PROGRAM main
  VAR
    S1 AT %IX0.0  : BOOL; (* abrir, NA *)
    S2 AT %IX0.1  : BOOL; (* cerrar, NA *)
    S0 AT %IX0.2  : BOOL; (* parada, NC: TRUE sin pulsar *)
    B1 AT %IX0.3  : BOOL; (* final: portón abierto *)
    B2 AT %IX0.4  : BOOL; (* final: portón cerrado *)
    B3 AT %IX0.5  : BOOL; (* barrera: obstáculo en el paso *)
    KM1 AT %QX0.0 : BOOL; (* motor: abrir *)
    KM2 AT %QX0.1 : BOOL; (* motor: cerrar *)
    H1 AT %QX0.2  : BOOL; (* baliza de movimiento *)
    ETAPA         : INT; (* 0 parado, 1 abriendo, 2 cerrando *)
    E0            : BOOL; (* ETAPA = 0 *)
    E1            : BOOL; (* ETAPA = 1 *)
    E2            : BOOL; (* ETAPA = 2 *)
  END_VAR
  VAR  (* added by the conversion: wires and edge detectors of the diagram *)
    _EQ1_OUT : BOOL;
    _EQ5_OUT : BOOL;
    _EQ9_OUT : BOOL;
    _NOT17_OUT : BOOL;
    _AND14_OUT : BOOL;
    _SEL13_OUT : INT;
    _NOT26_OUT : BOOL;
    _AND23_OUT : BOOL;
    _SEL22_OUT : INT;
    _AND32_OUT : BOOL;
    _SEL31_OUT : INT;
    _AND39_OUT : BOOL;
    _SEL38_OUT : INT;
    _AND46_OUT : BOOL;
    _SEL45_OUT : INT;
    _NOT53_OUT : BOOL;
    _SEL52_OUT : INT;
    _NOT62_OUT : BOOL;
  END_VAR

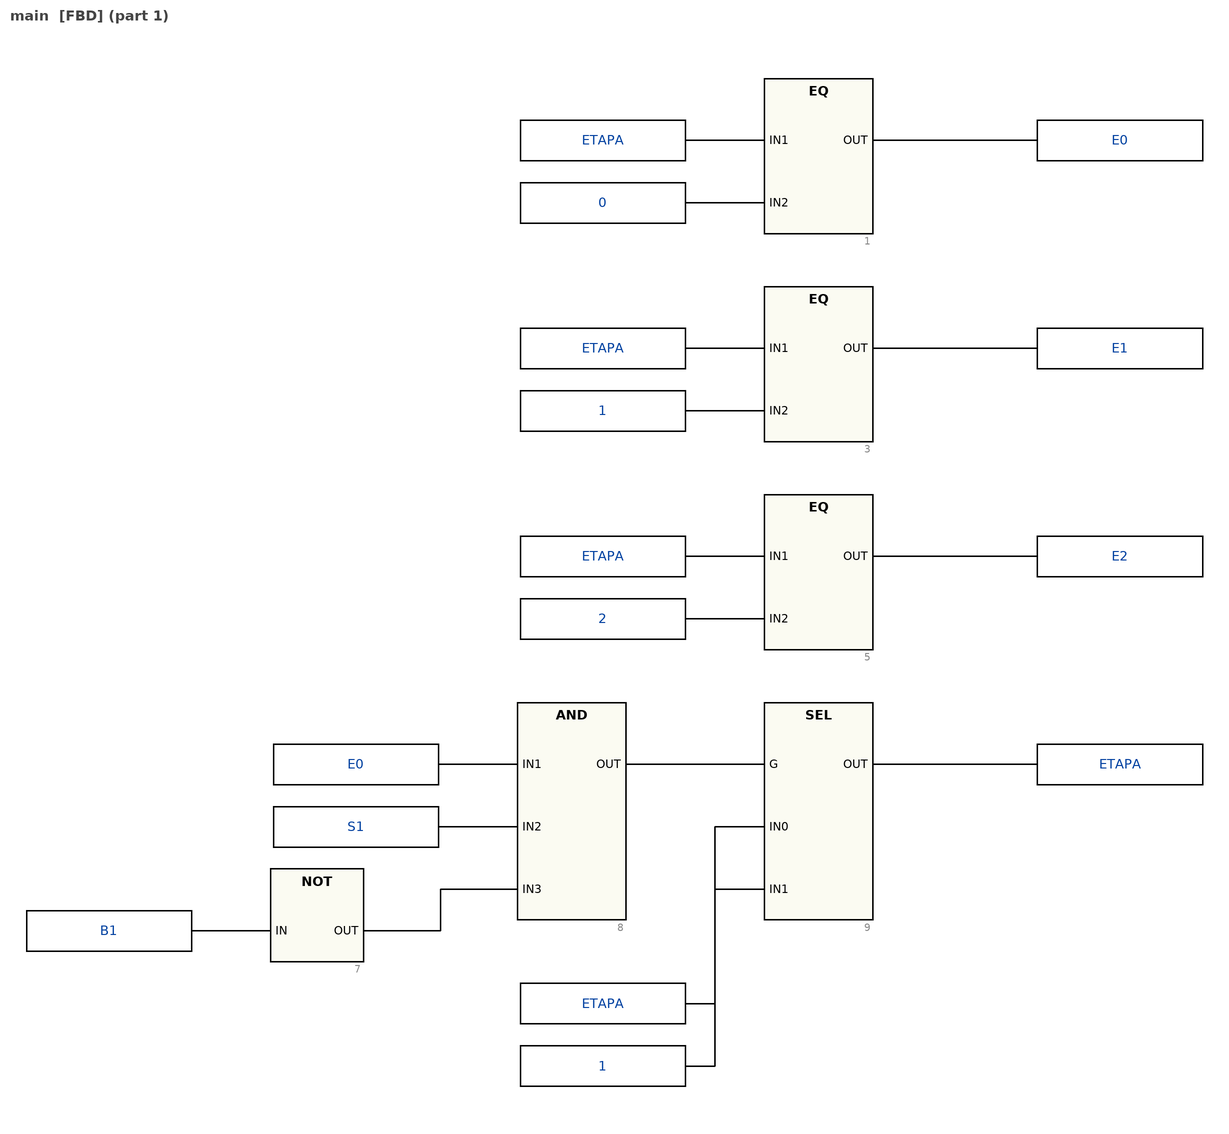
(* FBD diagram, written out as Structured Text *)
_EQ1_OUT := ETAPA = 0;
E0 := _EQ1_OUT;
_EQ5_OUT := ETAPA = 1;
E1 := _EQ5_OUT;
_EQ9_OUT := ETAPA = 2;
E2 := _EQ9_OUT;
_NOT17_OUT := NOT B1;
_AND14_OUT := E0 AND S1 AND _NOT17_OUT;
_SEL13_OUT := SEL(_AND14_OUT, ETAPA, 1);
ETAPA := _SEL13_OUT;
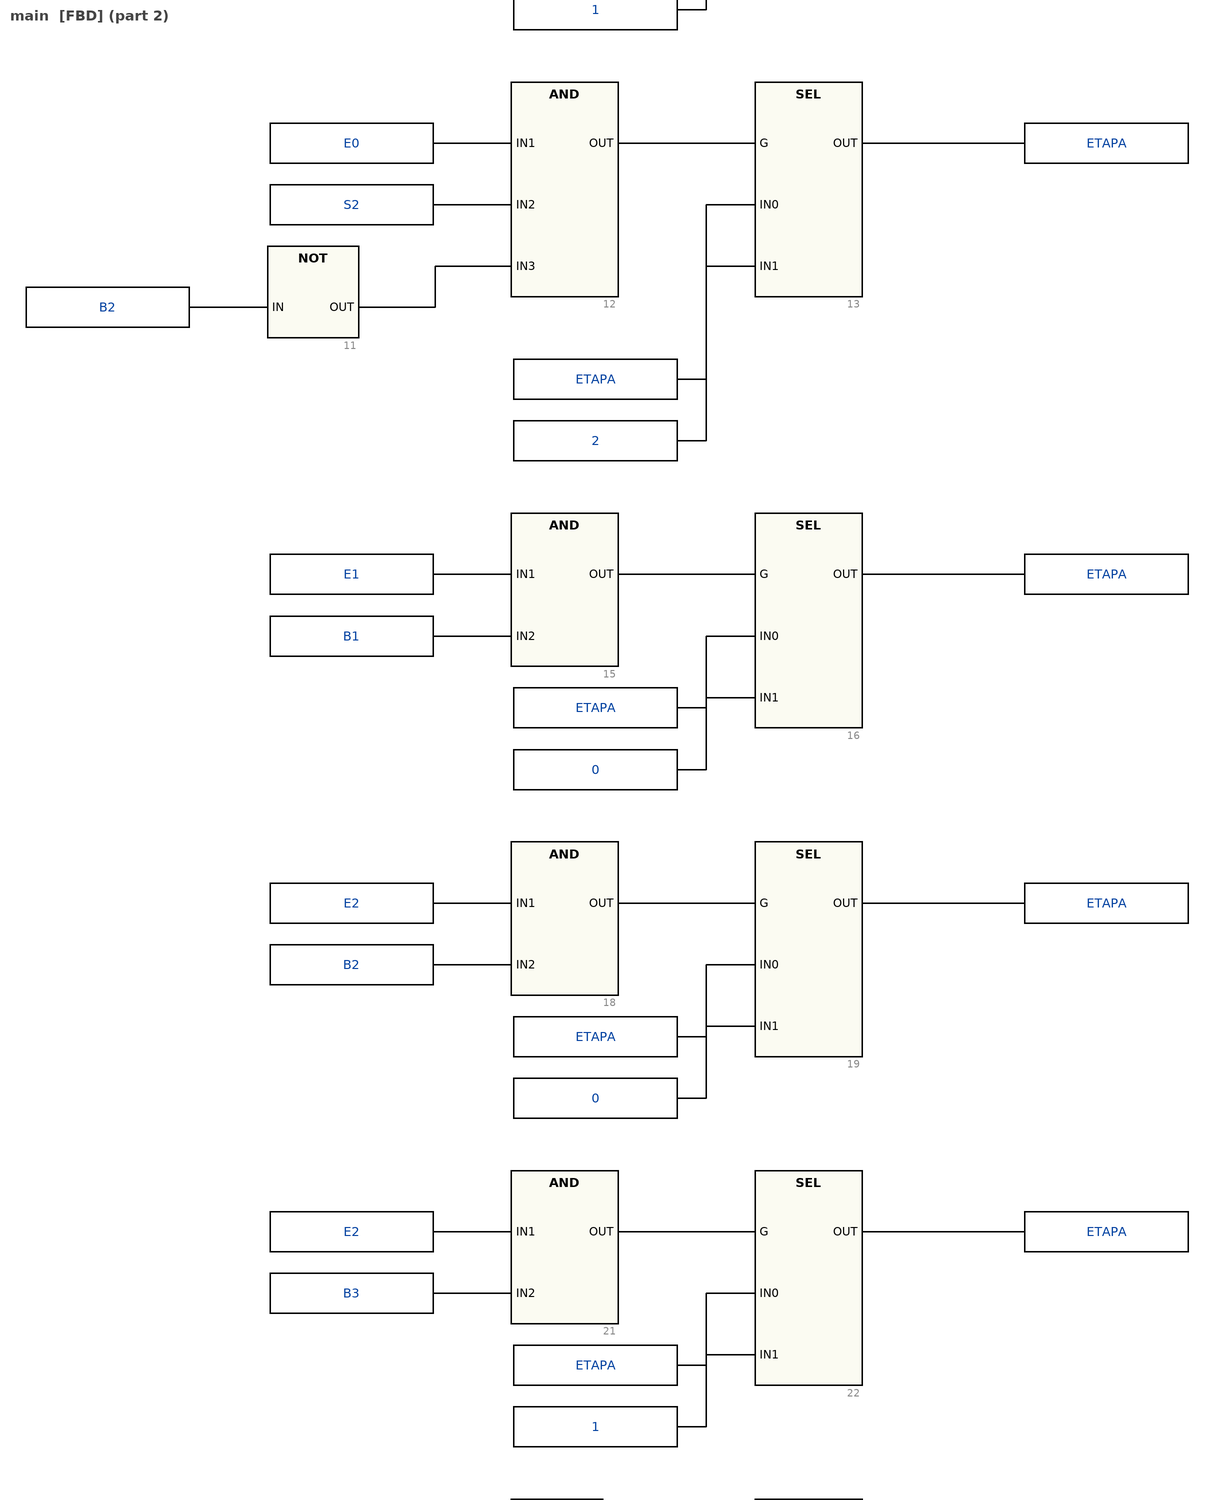
_NOT26_OUT := NOT B2;
_AND23_OUT := E0 AND S2 AND _NOT26_OUT;
_SEL22_OUT := SEL(_AND23_OUT, ETAPA, 2);
ETAPA := _SEL22_OUT;
_AND32_OUT := E1 AND B1;
_SEL31_OUT := SEL(_AND32_OUT, ETAPA, 0);
ETAPA := _SEL31_OUT;
_AND39_OUT := E2 AND B2;
_SEL38_OUT := SEL(_AND39_OUT, ETAPA, 0);
ETAPA := _SEL38_OUT;
_AND46_OUT := E2 AND B3;
_SEL45_OUT := SEL(_AND46_OUT, ETAPA, 1);
ETAPA := _SEL45_OUT;
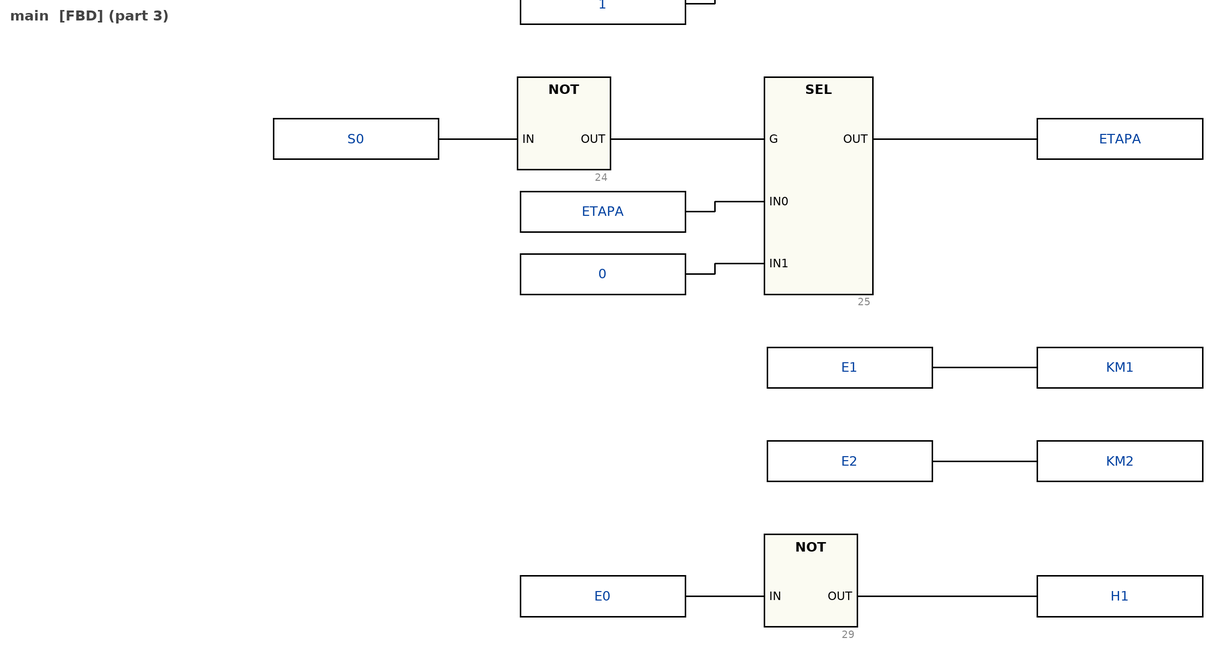
_NOT53_OUT := NOT S0;
_SEL52_OUT := SEL(_NOT53_OUT, ETAPA, 0);
ETAPA := _SEL52_OUT;
KM1 := E1;
KM2 := E2;
_NOT62_OUT := NOT E0;
H1 := _NOT62_OUT;
END_PROGRAM
